// TIA Portal V20 export
Screen "Pop-up_Hmi_Opmodes24_h_Popup"  740x540
  ScreenItem "Background" at 0,1 size 740x540  Type=HmiRectangle
  ScreenItem "Textfeld_1" at 74,100 size 34x38  Type=HmiTextBox
  ScreenItem "Text_HmiPanelNo" at 322,50 size 160x23  Type=HmiTextBox
  ScreenItem "State_OPMode8_Select" at 293,80 size 25x25  Type=HmiTextBox
  ScreenItem "State_OPMode8_NotSelect" at 293,80 size 25x25  Type=HmiTextBox
  ScreenItem "Descr_OPMode" at 174,26 size 305x20  Type=HmiTextBox
  ScreenItem "Overview_OPMode" at 1,1 size 657x25  Type=HmiTextBox
  ScreenItem "State_OPMode1_Select" at 111,80 size 25x25  Type=HmiTextBox
  ScreenItem "State_OPMode1_NotSelect" at 111,80 size 25x25  Type=HmiTextBox
  ScreenItem "State_OPMode2_Select" at 137,80 size 25x25  Type=HmiTextBox
  ScreenItem "State_OPMode2_NotSelect" at 137,80 size 25x25  Type=HmiTextBox
  ScreenItem "State_OPMode3_Select" at 163,80 size 25x25  Type=HmiTextBox
  ScreenItem "State_OPMode3_NotSelect" at 163,80 size 25x25  Type=HmiTextBox
  ScreenItem "State_OPMode4_Select" at 189,80 size 25x25  Type=HmiTextBox
  ScreenItem "State_OPMode4_NotSelect" at 189,80 size 25x25  Type=HmiTextBox
  ScreenItem "State_OPMode5_Select" at 215,80 size 25x25  Type=HmiTextBox
  ScreenItem "State_OPMode5_NotSelect" at 215,80 size 25x25  Type=HmiTextBox
  ScreenItem "State_OPMode6_Select" at 241,80 size 25x25  Type=HmiTextBox
  ScreenItem "State_OPMode6_NotSelect" at 241,80 size 25x25  Type=HmiTextBox
  ScreenItem "State_OPMode7_Select" at 267,80 size 25x25  Type=HmiTextBox
  ScreenItem "State_OPMode7_NotSelect" at 267,80 size 25x25  Type=HmiTextBox
  ScreenItem "State_OPMode9_Select" at 319,80 size 25x25  Type=HmiTextBox
  ScreenItem "State_OPMode9_NotSelect" at 319,80 size 25x25  Type=HmiTextBox
  ScreenItem "State_OPMode10_Select" at 345,80 size 25x25  Type=HmiTextBox
  ScreenItem "State_OPMode10_NotSelect" at 345,80 size 25x25  Type=HmiTextBox
  ScreenItem "State_OPMode11_Select" at 371,80 size 25x25  Type=HmiTextBox
  ScreenItem "State_OPMode11_NotSelect" at 371,80 size 25x25  Type=HmiTextBox
  ScreenItem "State_OPMode12_Select" at 397,80 size 25x25  Type=HmiTextBox
  ScreenItem "State_OPMode12_NotSelect" at 397,80 size 25x25  Type=HmiTextBox
  ScreenItem "State_OPMode13_Select" at 424,80 size 25x25  Type=HmiTextBox
  ScreenItem "State_OPMode13_NotSelect" at 424,80 size 25x25  Type=HmiTextBox
  ScreenItem "State_OPMode14_Select" at 450,80 size 25x25  Type=HmiTextBox
  ScreenItem "State_OPMode14_NotSelect" at 450,80 size 25x25  Type=HmiTextBox
  ScreenItem "State_OPMode15_Select" at 476,80 size 25x25  Type=HmiTextBox
  ScreenItem "State_OPMode15_NotSelect" at 476,80 size 25x25  Type=HmiTextBox
  ScreenItem "State_OPMode16_Select" at 502,80 size 25x25  Type=HmiTextBox
  ScreenItem "State_OPMode16_NotSelect" at 502,80 size 25x25  Type=HmiTextBox
  ScreenItem "State_OPMode17_Select" at 528,80 size 25x25  Type=HmiTextBox
  ScreenItem "State_OPMode17_NotSelect" at 528,80 size 25x25  Type=HmiTextBox
  ScreenItem "State_OPMode18_Select" at 554,80 size 25x25  Type=HmiTextBox
  ScreenItem "State_OPMode18_NotSelect" at 554,80 size 25x25  Type=HmiTextBox
  ScreenItem "State_OPMode19_Select" at 580,80 size 25x25  Type=HmiTextBox
  ScreenItem "State_OPMode19_NotSelect" at 580,80 size 25x25  Type=HmiTextBox
  ScreenItem "State_OPMode20_Select" at 606,80 size 25x25  Type=HmiTextBox
  ScreenItem "State_OPMode20_NotSelect" at 606,80 size 25x25  Type=HmiTextBox
  ScreenItem "State_OPMode21_Select" at 632,80 size 25x25  Type=HmiTextBox
  ScreenItem "State_OPMode21_NotSelect" at 632,80 size 25x25  Type=HmiTextBox
  ScreenItem "State_OPMode22_Select" at 658,80 size 25x25  Type=HmiTextBox
  ScreenItem "State_OPMode22_NotSelect" at 658,80 size 25x25  Type=HmiTextBox
  ScreenItem "State_OPMode23_Select" at 684,80 size 25x25  Type=HmiTextBox
  ScreenItem "State_OPMode23_NotSelect" at 684,80 size 25x25  Type=HmiTextBox
  ScreenItem "State_OPMode24_Select" at 710,80 size 25x25  Type=HmiTextBox
  ScreenItem "State_OPMode24_NotSelect" at 710,80 size 25x25  Type=HmiTextBox
  ScreenItem "Button_Back" at 1,1 size 90x60  Type=HmiButton
  ScreenItem "Button_Close" at 647,0 size 90x60  Type=HmiButton
  ScreenItem "Text_OPModeArea" at -84,288 size 260x25  Type=HmiTextBox
  ScreenItem "State_OPMode8_Vis" at 182,0 size 25x25  Type=HmiRectangle
  ScreenItem "State_OPMode1_Vis" at 0,0 size 25x25  Type=HmiRectangle
  ScreenItem "State_OPMode2_Vis" at 26,0 size 25x25  Type=HmiRectangle
  ScreenItem "State_OPMode3_Vis" at 52,0 size 25x25  Type=HmiRectangle
  ScreenItem "State_OPMode4_Vis" at 78,0 size 25x25  Type=HmiRectangle
  ScreenItem "State_OPMode5_Vis" at 104,0 size 25x25  Type=HmiRectangle
  ScreenItem "State_OPMode6_Vis" at 130,0 size 25x25  Type=HmiRectangle
  ScreenItem "State_OPMode7_Vis" at 156,0 size 25x25  Type=HmiRectangle
  ScreenItem "State_OPMode9_Vis" at 208,0 size 25x25  Type=HmiRectangle
  ScreenItem "State_OPMode10_Vis" at 234,0 size 25x25  Type=HmiRectangle
  ScreenItem "State_OPMode11_Vis" at 260,0 size 25x25  Type=HmiRectangle
  ScreenItem "State_OPMode12_Vis" at 286,0 size 25x25  Type=HmiRectangle
  ScreenItem "State_OPMode13_Vis" at 313,0 size 25x25  Type=HmiRectangle
  ScreenItem "State_OPMode14_Vis" at 339,0 size 25x25  Type=HmiRectangle
  ScreenItem "State_OPMode15_Vis" at 365,0 size 25x25  Type=HmiRectangle
  ScreenItem "State_OPMode16_Vis" at 391,0 size 25x25  Type=HmiRectangle
  ScreenItem "State_OPMode17_Vis" at 417,0 size 25x25  Type=HmiRectangle
  ScreenItem "State_OPMode18_Vis" at 443,0 size 25x25  Type=HmiRectangle
  ScreenItem "State_OPMode19_Vis" at 469,0 size 25x25  Type=HmiRectangle
  ScreenItem "State_OPMode20_Vis" at 495,0 size 25x25  Type=HmiRectangle
  ScreenItem "State_OPMode21_Vis" at 521,0 size 25x25  Type=HmiRectangle
  ScreenItem "State_OPMode22_Vis" at 547,0 size 25x25  Type=HmiRectangle
  ScreenItem "State_OPMode23_Vis" at 573,0 size 25x25  Type=HmiRectangle
  ScreenItem "State_OPMode24_Vis" at 599,0 size 25x25  Type=HmiRectangle
